// LS Electric XG5000 project: R10
// PLC LSPLC

PROGRAM NewProgram (task: 스캔 프로그램)

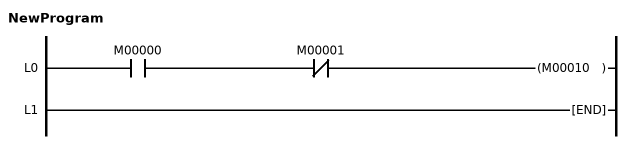
; L0
LOAD      M00000
AND NOT   M00001
OUT       M00010
; L1
END